Staubli VAL3: waitLoad.pgx

public program waitLoad(num x_nLib)
  local string l_sPath
  local string l_sPath1
begin
  l_sPath="Disk://data/CustomerLib/lib"+toString("",x_nLib)+"/savePROG"

  do
    l_sPath1=progTemp:libPath()
    delay(0)
  until l_sPath==l_sPath1
end
